(* IEC 61131-3 sources: FACTORY_io/fabrica-viva/etapa-2, 3 files *)

(* ---- fragmento-bloques.st ---- *)
(* ===== Etapa 2 · Bloque de función FB_Cinta =====
   Una cinta con vigilancia de atasco, para usar una instancia por cinta. Complétalo:
   - Motor sigue a Habilitar, salvo cuando hay Atasco.
   - Atasco se activa si Presencia lleva 3 s seguidos a TRUE con el motor en marcha (una caja parada
     delante de la fotocélula) y se queda activo hasta Rearme. *)
FUNCTION_BLOCK FB_Cinta
VAR_INPUT
  Habilitar : BOOL;   (* la cinta debe moverse *)
  Presencia : BOOL;   (* la fotocélula de vigilancia de esta cinta *)
  Rearme : BOOL;      (* borra el atasco *)
END_VAR
VAR_OUTPUT
  Motor : BOOL;       (* orden al motor de la cinta *)
  Atasco : BOOL;      (* atasco detectado, con memoria hasta Rearme *)
END_VAR
VAR
  (* tus variables internas del bloque *)
END_VAR

(* ---- tu código del bloque ---- *)
END_FUNCTION_BLOCK

(* ---- solucion.st ---- *)
(* Fábrica viva · Etapa 2 · Solución de referencia: FB_Cinta reutilizable, atasco que para toda la
   línea y rechazo de cajas sin etiqueta. *)
FUNCTION_BLOCK FB_Cinta
VAR_INPUT
  Habilitar : BOOL;
  Presencia : BOOL;
  Rearme : BOOL;
END_VAR
VAR_OUTPUT
  Motor : BOOL;
  Atasco : BOOL;
END_VAR
VAR
  Tapada : TON;
END_VAR

(* Solo cuenta con el motor en marcha: una caja delante de la fotocélula con la cinta parada no es un atasco. *)
Tapada(IN := Presencia AND Motor, PT := T#3s);
IF Rearme THEN
  Atasco := FALSE;
END_IF;
IF Tapada.Q THEN
  Atasco := TRUE;
END_IF;
Motor := Habilitar AND NOT Atasco;
END_FUNCTION_BLOCK

VAR_INPUT
  Marcha : BOOL;
  Paro : BOOL;
  Seta : BOOL;
  FotocelulaRecepcion : BOOL;
  CajasRecibidas : INT;
END_VAR
VAR_OUTPUT
  CintaRecepcion : BOOL;
  Alimentador : BOOL;
  Baliza : INT;
END_VAR
VAR
  EnMarcha : BOOL;
END_VAR

VAR_INPUT
  Rearme : BOOL;
  FotocelulaAtasco : BOOL;
  LecturaOk : BOOL;
  CodigoCaja : DINT;
  FotocelulaRechazo : BOOL;
  CajasRechazadas : INT;
  CajasFinLinea : INT;
END_VAR
VAR_OUTPUT
  CintaControl : BOOL;
  Desvio : BOOL;
  AlarmaAtasco : BOOL;
END_VAR
VAR
  Control : FB_Cinta;
  Leida : R_TRIG;
  Llega : R_TRIG;
  SinEtiqueta : BOOL;
  Pendiente : BOOL;
  Retardo : TON;
  Empuje : TP;
END_VAR

(* Etapa 1, retocada: el atasco también corta la marcha de toda la línea. *)
EnMarcha := (Marcha OR EnMarcha) AND NOT Paro AND Seta AND NOT AlarmaAtasco;
CintaRecepcion := EnMarcha;
Alimentador := EnMarcha;

(* Etapa 2: la cinta de control con su vigilancia. *)
Control(Habilitar := EnMarcha, Presencia := FotocelulaAtasco, Rearme := Rearme);
CintaControl := Control.Motor;
AlarmaAtasco := Control.Atasco;

(* Baliza: emergencia, atasco, marcha o parada. *)
IF NOT Seta THEN
  Baliza := 4;
ELSIF AlarmaAtasco THEN
  Baliza := 6;
ELSIF EnMarcha THEN
  Baliza := 1;
ELSE
  Baliza := 2;
END_IF;

(* Rechazo: el lector dice si la caja que entra lleva etiqueta; se aparta al llegar al desvío. *)
Leida(CLK := LecturaOk);
IF Leida.Q THEN
  SinEtiqueta := CodigoCaja = 0;
END_IF;
Llega(CLK := FotocelulaRechazo);
IF Llega.Q AND SinEtiqueta AND EnMarcha THEN
  Pendiente := TRUE;
END_IF;
Retardo(IN := Pendiente, PT := T#450ms);
IF Retardo.Q OR NOT EnMarcha THEN
  Pendiente := FALSE;
END_IF;
Empuje(IN := Retardo.Q, PT := T#600ms);
Desvio := Empuje.Q AND EnMarcha;

(* ---- fragmento-declaraciones.st ---- *)
(* ===== Etapa 2 · Control de entrada: señales nuevas ===== *)
VAR_INPUT
  Rearme : BOOL;              (* pulsador de rearme de la zona de control *)
  FotocelulaAtasco : BOOL;    (* vigilancia de atasco al principio de la cinta de control *)
  LecturaOk : BOOL;           (* el lector de códigos: pulso al leer una caja *)
  CodigoCaja : DINT;          (* el código leído; 0 = caja sin etiqueta *)
  FotocelulaRechazo : BOOL;   (* fotocélula justo antes del desvío de rechazo *)
  CajasRechazadas : INT;      (* cajas retiradas en la cinta de rechazo *)
  CajasFinLinea : INT;        (* cajas que llegan al final de la línea *)
END_VAR
VAR_OUTPUT
  CintaControl : BOOL;        (* la cinta de control y la de rechazo *)
  Desvio : BOOL;              (* el empujador de rechazo *)
  AlarmaAtasco : BOOL;        (* hay un atasco en la zona de control *)
END_VAR
VAR
  Control : FB_Cinta;         (* la cinta de control, vigilada por tu bloque *)
END_VAR
